FUNCTION_BLOCK FallbackElapsedTime (* Composite Function Block Type *)
  (* Standard: 61499-2 *)
  (* Version 0.0, 10/7/2026, Schneider Electric, template *)
  PACKAGE SE.Nereda;
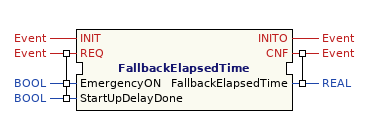
  EVENT_INPUT
    INIT; (* Initialization Request *)
    REQ WITH EmergencyON, StartUpDelayDone; (* Normal Execution Request *)
  END_EVENT
  EVENT_OUTPUT
    INITO; (* Initialization Confirm *)
    CNF WITH FallbackElapsedTime; (* Execution Confirmation *)
  END_EVENT
  VAR_INPUT
    EmergencyON : BOOL; (* Input event qualifier *)
    StartUpDelayDone : BOOL; (* Input event qualifier *)
  END_VAR
  VAR_OUTPUT
    FallbackElapsedTime : REAL; (* Output event qualifier *)
  END_VAR
  FBS
    FallbackElapsedTimeCalc : devMntCalc(TBaseOperationDuration := T#1s, TBaseElapsedDuration := T#1d); {SET_ATTRIBUTE(Configuration.Component.HideUnusedPorts, )}
    FB1 : UDINT2REAL;
    FB2 : BOOL2INT;
    FB3 : AND_88A3DD8EC65DD11C; {SET_ATTRIBUTE(Configuration.GenericFBType.InterfaceParams, Runtime.Standard#CNT:=2;OUT:BOOL)}
    FB4 : DIVIDE(pin_02E479D09E2C7EA2 := 60);
  END_FBS
  EVENT_CONNECTIONS
    INIT TO FallbackElapsedTimeCalc.INIT;
    FallbackElapsedTimeCalc.INITO TO INITO;
    FallbackElapsedTimeCalc.CNF_OPD TO FB1.DD5870AA881150BB;
    REQ TO FB3.REQ;
    FB2.6FC99A5BD1C38561 TO FallbackElapsedTimeCalc.REQ_PV;
    FB1.6FC99A5BD1C38561 TO FB4.0FDF8A587C3CA146;
    FB3.CNF TO FB2.DD5870AA881150BB;
    FB4.6D05A744943B688E TO CNF;
  END_CONNECTIONS
  DATA_CONNECTIONS
    FallbackElapsedTimeCalc.CurrentOperationDuration TO FB1.4573FC8F228EB71D;
    EmergencyON TO FB3.IN1;
    FB2.A6DEF5F9C27C1848 TO FallbackElapsedTimeCalc.Pv;
    FB1.A6DEF5F9C27C1848 TO FB4.8EF5C40F2FEA5451;
    StartUpDelayDone TO FB3.IN2;
    FB3.OUT TO FB2.4573FC8F228EB71D;
    FB4.E78A8A65D4120686 TO FallbackElapsedTime;
  END_CONNECTIONS
END_FUNCTION_BLOCK
